(* PLC project PR_ModeManageNoMode_PLC, SiemensToBackhoff Siemens TIA Portal to Beckhoff TwinCAT PLCopen Converter 2.0 *)
(* stored: creationDateTime 2026-09-28T10:47:49.957897, modificationDateTime 2026-09-28T10:47:49.957897 *)

FUNCTION_BLOCK PR_ModeManageNoMode
VAR_INPUT
	iFirstscan : BOOL;  // PLC First Scan Bit
	iControlOn : BOOL;  // Machine All Safety Relay Healthy
	iAutoModeEnable : BOOL;  // If conditions are OK to start automode make this bit high
	iManModeEnable : BOOL;  // If conditions are OK to sart manual mode make this bit high
	iAutoMode : BOOL;  // Auto Mode Input PB/SW
	iManMode : BOOL;  // Man Mode Input PB/SW
	iCycleStart : BOOL;  // Cycle Start Input PB
	iCycleStop : BOOL;  // Cycle Stop Input PB (NC Type)
	iHomePB : BOOL;  // Home Input PB
	iEndOfCycle : BOOL;  // If Cycle Completed make this bit high
	iDrainCycle : BOOL;  // If conditions are OK to start drain cycle make this bit high
	iDryCycle : BOOL;  // If conditions are OK to start dry cycle make this bit high
	iDrainCompleted : BOOL;  // If Drain Completed make this bit high
	iHomeCompleted : BOOL;  // If Home Completed make this bit high
	iImmediateStop : BOOL;  // To abort autocycle or to select manual while running in auto make this bit 1
	iCycleStartDelay : TIME;  // Cycle Start PB Press Delay Eg. If 2Sec T#2S
	iBypassHomeOption : BOOL;  // Make sure that autocycle can initiate without home condition = 1
END_VAR
VAR_OUTPUT
	qManModeActive : BOOL;  // Man Mode Active
	qWaitForCStart : BOOL;  // Waiting For Cycle Start
	qAutoRunningActive : BOOL;  // AutoRunning Active
	qHomeRunningActive : BOOL;  // Home Running Active
	qDrainActive : BOOL;  // Drain Active
	qCycleStopActive : BOOL;  // Cycle Stop Active
	qDryCycleActive : BOOL;  // Dry Cycle Active
	qModuleReset : BOOL;  // 1 If No Mode Selected
	qMsgCStartandNoHome : BOOL;  // Cycle Start PB Pressed but MC Not at Home
	qMsgManModeinAutoRunning : BOOL;  // Manual Mode selected during Auto Running
END_VAR
VAR
	sPowerOnReset : BOOL;  // Power ON reset Bit during initial power ON
	sControlOnPulse : BOOL;  // Control ON pulse
	sControlOnEdge : R_TRIG;  // Control ON Input Positive Edge
	sManModeActivePulse : R_TRIG;  // Man Mode Active Positive Edge Pulse
	sCycleStartDelay : TIME;  // Cycle Start Delay
	CycleStartOnDelayTimer : TON;  // ON Delay Timer SFB4
	sAutoRunningActive : BOOL;  // Auto Running Active
	sManModeActive : BOOL;  // Man Mode Active
	sHomeRunningActive : BOOL;  // Home Running Active
	sWaitForCStart : BOOL;  // Waiting For Cycle Start
	sDrainActive : BOOL;  // Drain Active
	sDryCycleActive : BOOL;  // Dry Cycle Active
	sCycleStopActive : BOOL;  // Cycle Stop Active
	sModuleReset : BOOL;  // Module Reset
	sMsgCStartandNoHome : BOOL;  // Cycle Start PB Pressed but MC Not at Home
	sMsgManModeinAutoRunning : BOOL;  // Manual Mode selected during Auto Running
END_VAR
  VAR  (* added by the conversion: wires and edge detectors of the diagram *)
    _GT8_ENO : BOOL;
    _GT8_OUT : BOOL;
    _LT11_ENO : BOOL;
    _LT11_OUT : BOOL;
  END_VAR

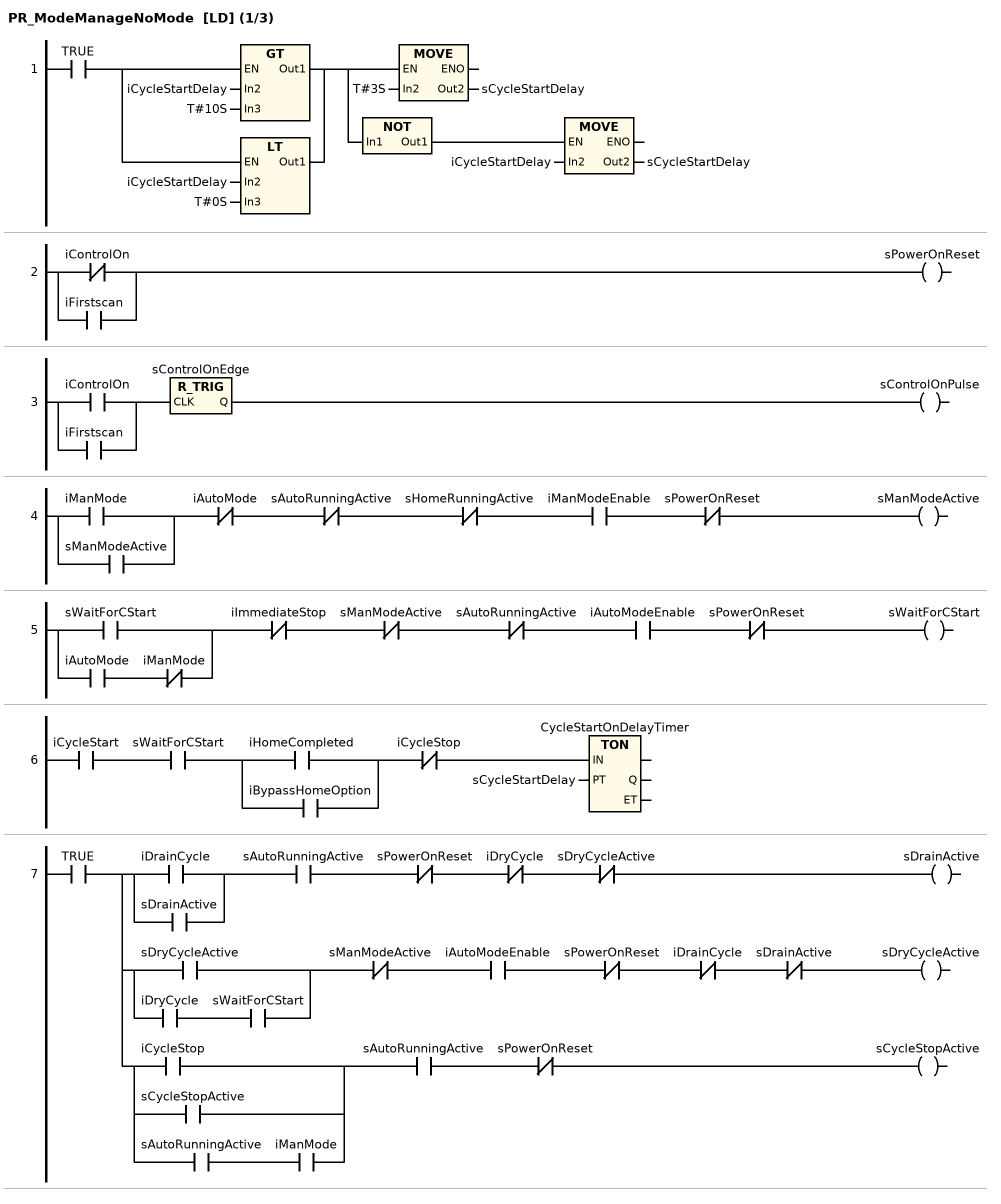
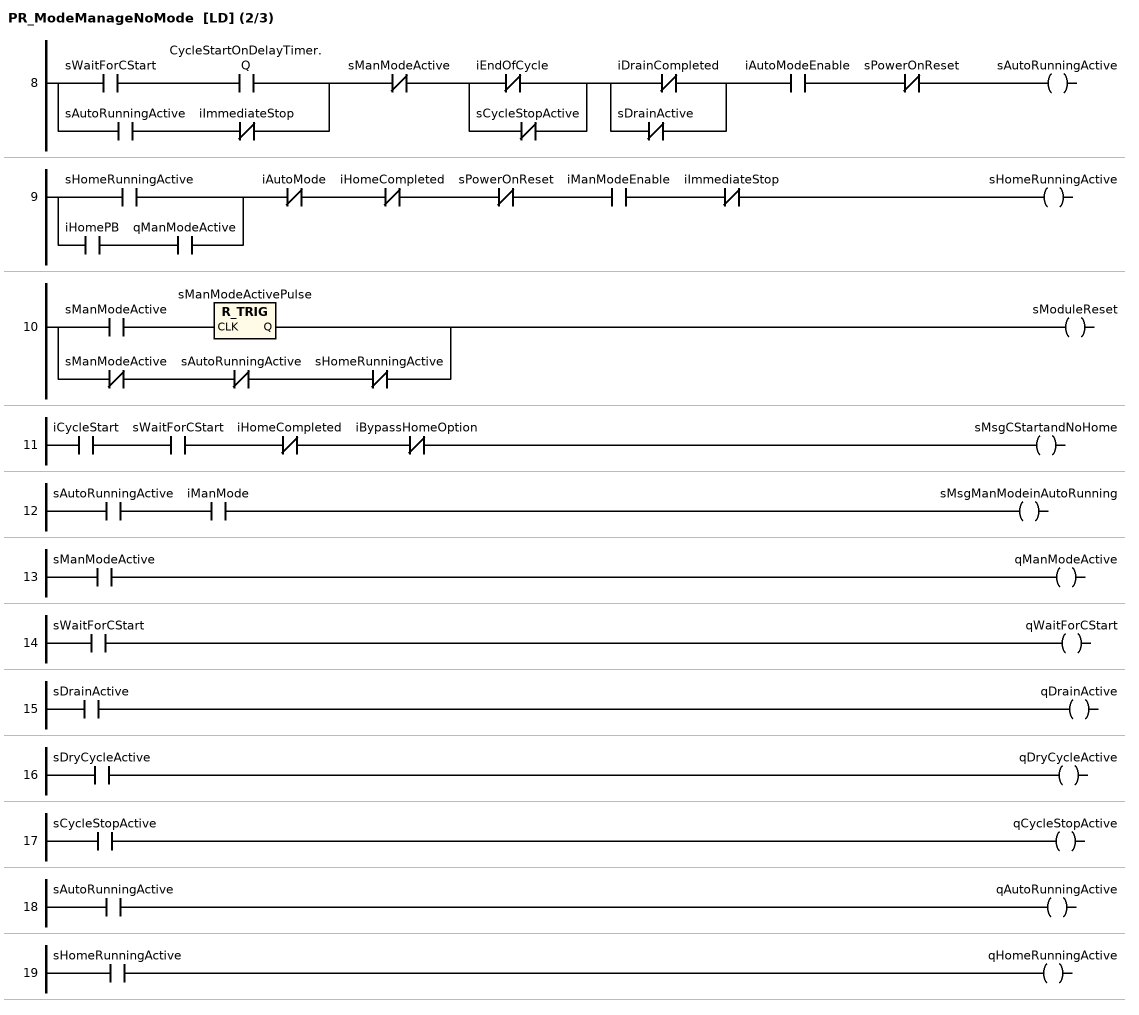
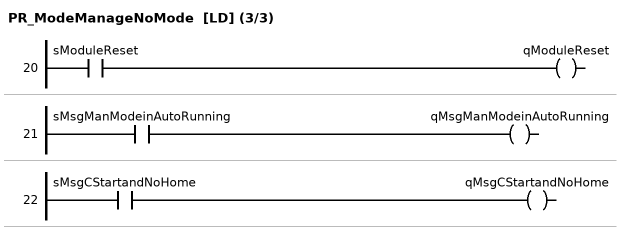
(* LD diagram, written out as Structured Text *)
(* ==============================================================================
 Company: Precision Automation & Robotics India Ltd. 
------------------------------------------------------------------------------
 Item Code: S11002022002
 Author/Created by: PARI
 Reviewed/Checked by: Atul P
 First Release on: 14-Aug-2015
 Latest update on: 14-Aug-2015
------------------------------------------------------------------------------
 Tested with: CPU firmware, model or simulator testing
 Engineering/Editor: TIA Portal V15.1
------------------------------------------------------------------------------
 Restrictions: No
 Dependencies/Requirements:
------------------------------------------------------------------------------
 Change Log:
 Ver.	Date		Changed by		Details of changes
 1.0       14-Aug-2015                           A.D	                                     First release version
------------------------------------------------------------------------------
Functionality:
This block is used Control Mode Of System.After Power On or End Of Cycle It 
will go to No Mode State if mode 
Selection is not present

 Inputs
iFirstscan	Bool
iContolOn	Bool
iAutoModeEnable	Bool
iManModeEnable	Bool
iAutoMode	Bool
iManMode	Bool
iCycleStart	Bool
iCycleStop	Bool
iHomePB	Bool
iEndOfCycle	Bool
iDrainCycle	Bool
iDryCycle	Bool
iDrainCompleted	Bool
iHomeCompleted	Bool
iImmediateStop	Bool
iCycleStartDelay	Time
iBypassHomeOption	Bool


 Outputs
qManModeActive	Bool
qWaitForCStart	Bool
qAutoRunningActive	Bool
qHomeRunningActive	Bool
qDrainActive	Bool
qCycleStopActive	Bool
qDryCycleActive	Bool
qModuleReset	Bool


In-outs
Nill

------------------------------------------------------------------------------
Errors reported:
Nill

Messages:
qMsgCStartandNoHome	Bool
qMsgManModeinAutoRunning	Bool

============================================================================== *)

(* Cycle Start delay validation *)

_GT8_OUT := GT(EN := TRUE, IN1 := iCycleStartDelay, IN2 := T#10S, ENO => _GT8_ENO);
_LT11_OUT := LT(EN := TRUE, IN1 := iCycleStartDelay, IN2 := T#0S, ENO => _LT11_ENO);
IF _LT11_OUT OR _GT8_OUT THEN sCycleStartDelay := T#3S; END_IF;
IF NOT (_LT11_OUT OR _GT8_OUT) THEN sCycleStartDelay := iCycleStartDelay; END_IF;
(* Power ON reset Bit during initial power ON
Reset Active *)

sPowerOnReset := NOT iControlOn OR iFirstscan;
(* Control On pulse
#sControlOnPulse *)

sControlOnEdge(CLK := iControlOn OR iFirstscan);
sControlOnPulse := sControlOnEdge.Q;
(* Manual mode active
Man Mode *)

sManModeActive := (iManMode OR sManModeActive) AND NOT iAutoMode AND NOT sAutoRunningActive AND NOT sHomeRunningActive AND iManModeEnable AND NOT sPowerOnReset;
(* Waiting for cycle to start
Auto Mode *)

sWaitForCStart := (iAutoMode AND NOT iManMode OR sWaitForCStart) AND NOT iImmediateStop AND NOT sManModeActive AND NOT sAutoRunningActive AND iAutoModeEnable AND NOT sPowerOnReset;
(* CycleStartDelayTimer *)

CycleStartOnDelayTimer(IN := iCycleStart AND sWaitForCStart AND (iHomeCompleted OR iBypassHomeOption) AND NOT iCycleStop, PT := sCycleStartDelay);
(* Drain,Dry,Cycle Stop Active *)

sDrainActive := TRUE AND (iDrainCycle OR sDrainActive) AND sAutoRunningActive AND NOT sPowerOnReset AND NOT iDryCycle AND NOT sDryCycleActive;
sDryCycleActive := TRUE AND (iDryCycle AND sWaitForCStart OR sDryCycleActive) AND NOT sManModeActive AND iAutoModeEnable AND NOT sPowerOnReset AND NOT iDrainCycle AND NOT sDrainActive;
sCycleStopActive := TRUE AND (iCycleStop OR sAutoRunningActive AND iManMode OR sCycleStopActive) AND sAutoRunningActive AND NOT sPowerOnReset;
(* Auto running active
Auto Running *)

sAutoRunningActive := (sWaitForCStart AND CycleStartOnDelayTimer.Q OR sAutoRunningActive AND NOT iImmediateStop) AND NOT sManModeActive AND (NOT iEndOfCycle OR NOT sCycleStopActive) AND (NOT iDrainCompleted OR NOT sDrainActive) AND iAutoModeEnable AND NOT sPowerOnReset;
(* Home running active *)

sHomeRunningActive := (iHomePB AND qManModeActive OR sHomeRunningActive) AND NOT iAutoMode AND NOT iHomeCompleted AND NOT sPowerOnReset AND iManModeEnable AND NOT iImmediateStop;
(* Resetting module to initial state
Module Reset *)

sManModeActivePulse(CLK := sManModeActive);
sModuleReset := NOT sManModeActive AND NOT sAutoRunningActive AND NOT sHomeRunningActive OR sManModeActivePulse.Q;
(* Message if machine is started without home conditions OK
Machine Not At Home if C Start Press *)

sMsgCStartandNoHome := iCycleStart AND sWaitForCStart AND NOT iHomeCompleted AND NOT iBypassHomeOption;
(* Message if manual mode selected during auto running
MsgManModeinAutoRunning *)

sMsgManModeinAutoRunning := sAutoRunningActive AND iManMode;
(* Outputs *)

qManModeActive := sManModeActive;
qWaitForCStart := sWaitForCStart;
qDrainActive := sDrainActive;
qDryCycleActive := sDryCycleActive;
qCycleStopActive := sCycleStopActive;
qAutoRunningActive := sAutoRunningActive;
qHomeRunningActive := sHomeRunningActive;
qModuleReset := sModuleReset;
qMsgManModeinAutoRunning := sMsgManModeinAutoRunning;
qMsgCStartandNoHome := sMsgCStartandNoHome;
END_FUNCTION_BLOCK
